PROGRAM main
  VAR
    button AT %QX0.0 : BOOL;
    Motor AT %QX0.1 : BOOL;
    Package_detected AT %QX0.2 : BOOL;
    reset AT %QX0.3 : BOOL;
    total_count AT %MW1 : INT;
    Big_Box AT %MW2 : INT;
    Medium_Box AT %MW3 : INT;
    small_box AT %MW4 : INT;
    is_small AT %MX0.0 : BOOL;
    is_BIG AT %MX0.1 : BOOL;
    weight AT %MW0 : INT;
    CTU0 : CTU;
    CTU1 : CTU;
    CTU_DINT0 : CTU_DINT;
    CTUD0 : CTUD;
    CTU2 : CTU;
    CTU3 : CTU;
  END_VAR

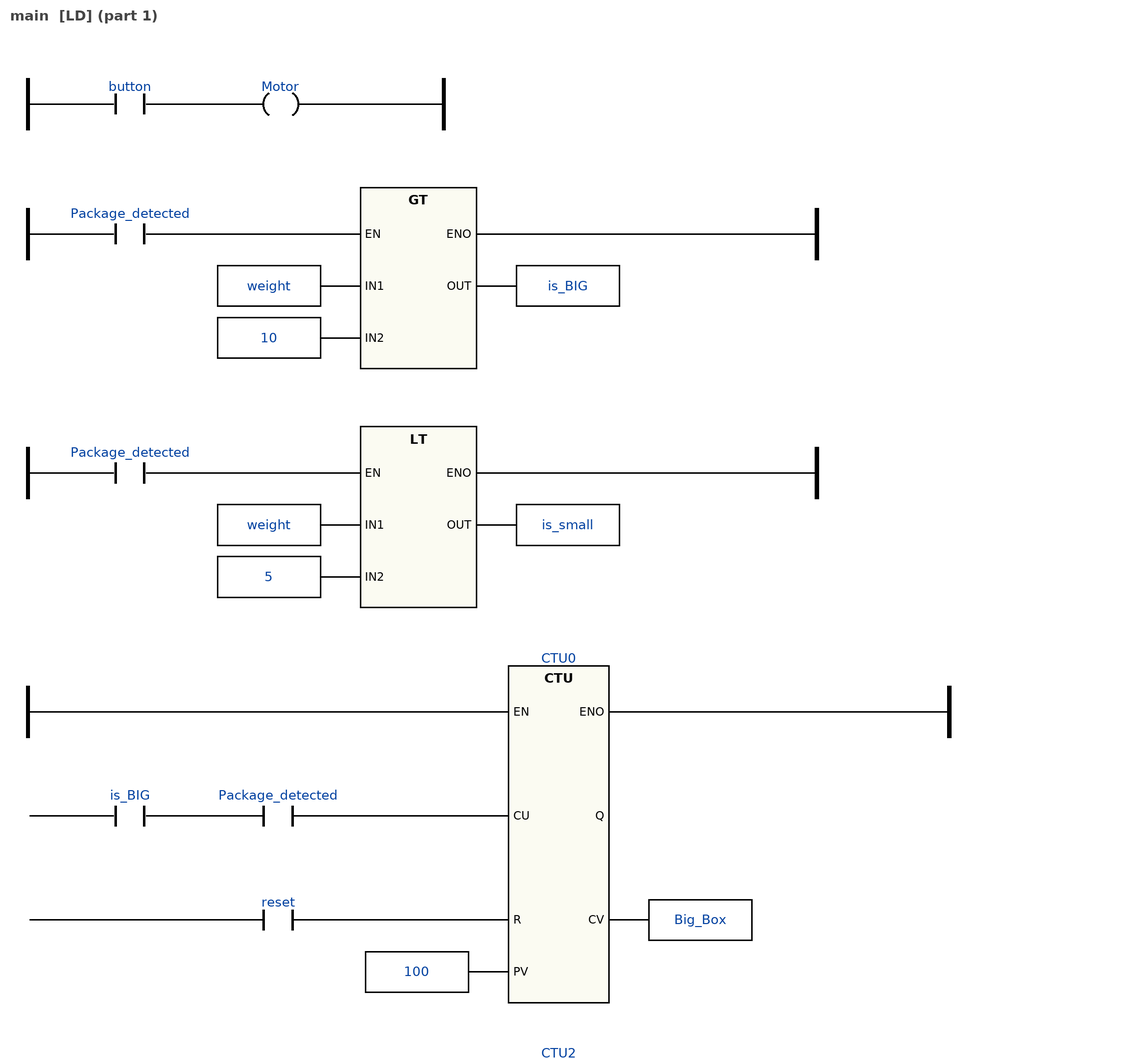
(* LD diagram, written out as Structured Text *)
Motor := button;
IF Package_detected THEN is_BIG := weight > 10; END_IF;
IF Package_detected THEN is_small := weight < 5; END_IF;
CTU0(CU := is_BIG AND Package_detected, R := reset, PV := 100);
Big_Box := CTU0.CV;
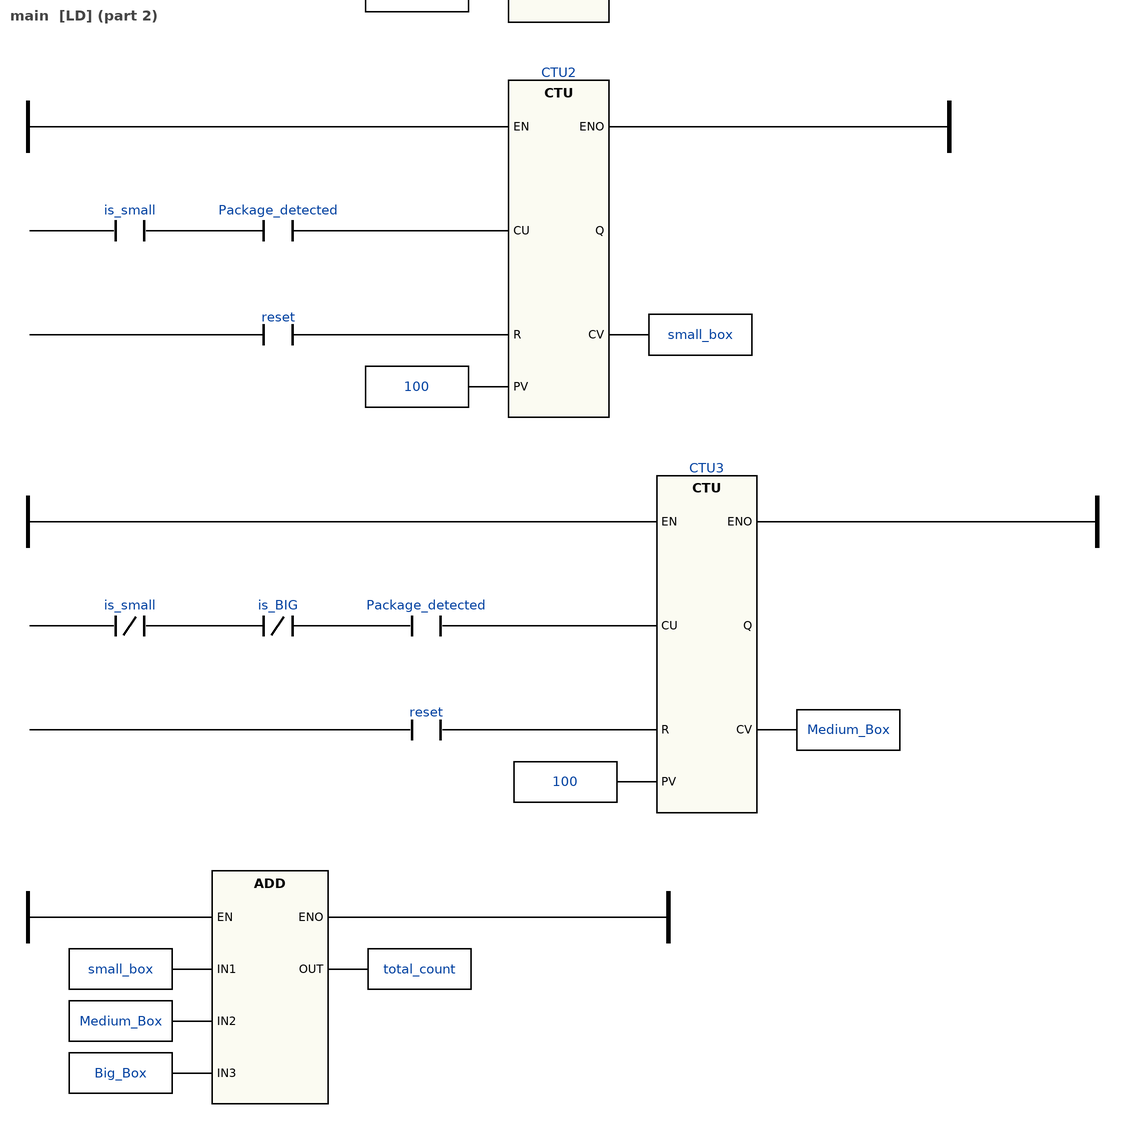
CTU2(CU := is_small AND Package_detected, R := reset, PV := 100);
small_box := CTU2.CV;
CTU3(CU := NOT is_small AND NOT is_BIG AND Package_detected, R := reset, PV := 100);
Medium_Box := CTU3.CV;
total_count := small_box + Medium_Box + Big_Box;
END_PROGRAM
